SUBAPPLICATION SoftKeySR_PC_A_OPC (* Geraet A (Station 11, 192.168.1.11): 2 SoftKeys (Set/Reset) rufen je einen eigenen argument- und rueckgabewertlosen OPC-UA-Methodenaufruf auf Geraet B auf (CLIENT_0, 2 eigene Methoden - wie Training_04, aber ohne Toggle); GreenWhiteBackground am Set-SoftKey zeigt den von Geraet B lokal ueberwachten Flipflop-Zustand - 'SUB style': das Protokoll steckt im MyLib::sys-Composite, nicht in der Resource des Geraets *)
  (* Standard: 61499-2; Description: Copyright (c) 2026 Meisterschulen am Ostbahnhof This program and the accompanying materials are made available under the terms of the Eclipse Public License 2.0 which is available at https://www.eclipse.org/legal/epl-2.0/ SPDX-License-Identifier: EPL-2.0 *)
  (* Version 1.0, 2026-09-03, Franz Höpfinger, Meisterschulen am Ostbahnhof, initial API and implementation and/or initial documentation *)
  PACKAGE MyLib::sys;
  IMPORT isobus::UT::Q::const::IDs::ID_NULL;
  IMPORT isobus::UT::io::Softkey::SoftKeyActivationCode::SK_RELEASED;
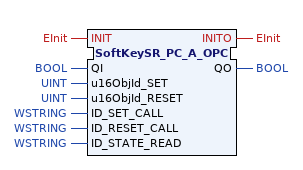
  EVENT_INPUT
    INIT : EInit; (* Initialization Request *)
  END_EVENT
  EVENT_OUTPUT
    INITO : EInit; (* Initialization Confirm *)
  END_EVENT
  VAR_INPUT
    QI : BOOL := TRUE; (* Quality Input - TRUE to enable service *)
    u16ObjId_SET : UINT := ID_NULL; (* Object ID SoftKey Set (traegt auch das GreenWhiteBackground) *)
    u16ObjId_RESET : UINT := ID_NULL; (* Object ID SoftKey Reset *)
    ID_SET_CALL : WSTRING; (* Remote-Methodenadresse (ACTION=CALL_METHOD) fuer den Set-Methodenaufruf auf Geraet B *)
    ID_RESET_CALL : WSTRING; (* Remote-Methodenadresse (ACTION=CALL_METHOD) fuer den Reset-Methodenaufruf auf Geraet B *)
    ID_STATE_READ : WSTRING; (* Lokal ueberwachte Adresse (BOOL, ACTION=READ) fuer den Flipflop-Zustand, wird von Geraet B remote beschrieben *)
  END_VAR
  VAR_OUTPUT
    QO : BOOL; (* Quality Output - TRUE if service executed successfully *)
  END_VAR
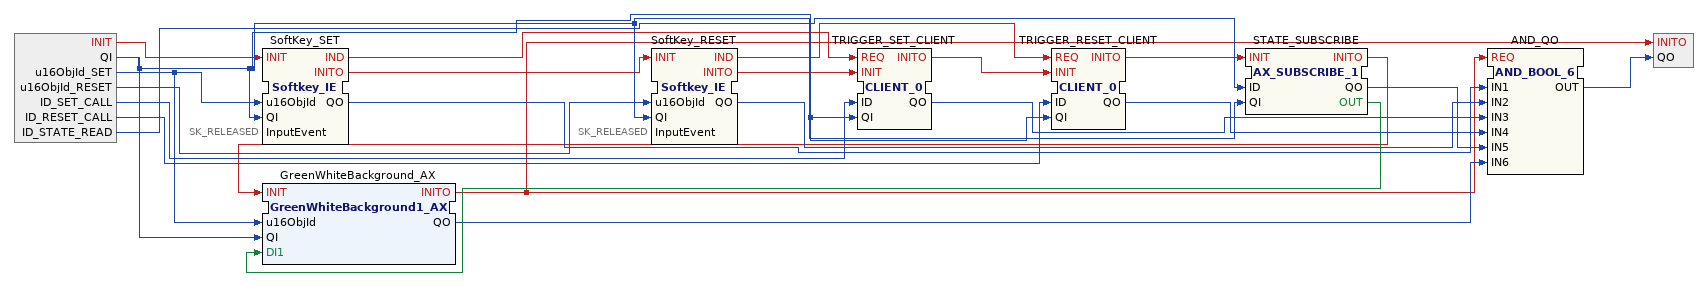
  FBS
    SoftKey_SET : isobus::UT::io::Softkey::Softkey_IE(InputEvent := SK_RELEASED);
    SoftKey_RESET : isobus::UT::io::Softkey::Softkey_IE(InputEvent := SK_RELEASED);
    TRIGGER_SET_CLIENT : iec61499::net::CLIENT_0;
    TRIGGER_RESET_CLIENT : iec61499::net::CLIENT_0;
    STATE_SUBSCRIBE : adapter::net::AX_SUBSCRIBE_1;
    AND_QO : iec61131::booleanOperators::AND_BOOL_6;
  END_FBS
  SUBAPPS
    GreenWhiteBackground_AX : MyLib::sys::GreenWhiteBackground1_AX;
  END_SUBAPPS
  EVENT_CONNECTIONS
    SoftKey_SET.IND TO TRIGGER_SET_CLIENT.REQ;
    SoftKey_RESET.IND TO TRIGGER_RESET_CLIENT.REQ;
    INIT TO SoftKey_SET.INIT;
    SoftKey_SET.INITO TO SoftKey_RESET.INIT;
    SoftKey_RESET.INITO TO TRIGGER_SET_CLIENT.INIT;
    TRIGGER_SET_CLIENT.INITO TO TRIGGER_RESET_CLIENT.INIT;
    TRIGGER_RESET_CLIENT.INITO TO STATE_SUBSCRIBE.INIT;
    STATE_SUBSCRIBE.INITO TO GreenWhiteBackground_AX.INIT;
    GreenWhiteBackground_AX.INITO TO INITO;
    GreenWhiteBackground_AX.INITO TO AND_QO.REQ;
  END_CONNECTIONS
  DATA_CONNECTIONS
    u16ObjId_SET TO SoftKey_SET.u16ObjId;
    u16ObjId_RESET TO SoftKey_RESET.u16ObjId;
    u16ObjId_SET TO GreenWhiteBackground_AX.u16ObjId;
    ID_SET_CALL TO TRIGGER_SET_CLIENT.ID;
    ID_RESET_CALL TO TRIGGER_RESET_CLIENT.ID;
    ID_STATE_READ TO STATE_SUBSCRIBE.ID;
    QI TO SoftKey_SET.QI;
    QI TO SoftKey_RESET.QI;
    QI TO TRIGGER_SET_CLIENT.QI;
    QI TO TRIGGER_RESET_CLIENT.QI;
    QI TO STATE_SUBSCRIBE.QI;
    SoftKey_SET.QO TO AND_QO.IN1;
    SoftKey_RESET.QO TO AND_QO.IN2;
    TRIGGER_SET_CLIENT.QO TO AND_QO.IN3;
    TRIGGER_RESET_CLIENT.QO TO AND_QO.IN4;
    STATE_SUBSCRIBE.QO TO AND_QO.IN5;
    AND_QO.OUT TO QO;
    QI TO GreenWhiteBackground_AX.QI;
    GreenWhiteBackground_AX.QO TO AND_QO.IN6;
  END_CONNECTIONS
  ADAPTER_CONNECTIONS
    STATE_SUBSCRIBE.OUT TO GreenWhiteBackground_AX.DI1;
  END_CONNECTIONS
END_SUBAPPLICATION
